(* IEC 61131-3 sources: genai_codesys/experiments/raw/formal/20261109_234635_2ba96d/public_02/custom__deepseek-v4.1-flash-1017/attempt_00, 2 files *)

(* ---- declaration.st ---- *)
FUNCTION_BLOCK FB_DWordEdgeDetection
VAR_INPUT
    value : DWORD;
END_VAR
VAR_OUTPUT
    hasChanged : BOOL;
    hasRisingEdges : BOOL;
    risingBits : DWORD;
    noOfRisingBits : USINT;
    hasFallingEdges : BOOL;
    fallingBits : DWORD;
    noOfFallingBits : USINT;
END_VAR
VAR
    previousValue : DWORD;
    countBits : DWORD;
    i : INT;
END_VAR

(* ---- implementation.st ---- *)
risingBits := value AND NOT previousValue;
fallingBits := (NOT value) AND previousValue;
hasChanged := value <> previousValue;
hasRisingEdges := risingBits <> DWORD#0;
hasFallingEdges := fallingBits <> DWORD#0;
noOfRisingBits := USINT#0;
countBits := risingBits;
FOR i := 0 TO 31 DO
    IF (countBits AND DWORD#1) <> DWORD#0 THEN
        noOfRisingBits := noOfRisingBits + USINT#1;
    END_IF;
    countBits := countBits / DWORD#2;
END_FOR;
noOfFallingBits := USINT#0;
countBits := fallingBits;
FOR i := 0 TO 31 DO
    IF (countBits AND DWORD#1) <> DWORD#0 THEN
        noOfFallingBits := noOfFallingBits + USINT#1;
    END_IF;
    countBits := countBits / DWORD#2;
END_FOR;
previousValue := value;
